(* IEC 61131-3 sources: sis-interlock-demo/src/DUTs/Sis, 21 files *)

(* ---- E_BypassState.dut.st ---- *)
// Назначение: состояние байпаса канала (диаграмма 5.7).
// Автор:      kr0nsch
// Версия:     0.1.0
// Документ:   docs/DESIGN.md, раздел «4.1 Перечисления»
// ВНИМАНИЕ:   код демонстрационный и не предназначен для систем безопасности. Реальная ПАЗ
//             требует определения SIL, сертифицированных аппаратных и программных средств
//             и валидации по ГОСТ Р МЭК 61511.
{attribute 'qualified_only'}
{attribute 'strict'}
TYPE E_BypassState :
(
    Off     := 0,    // байпаса нет
    Active  := 1,    // байпас действует, идёт отсчёт tBypassMax
    Expired := 2,    // срок истёк, запрос ещё держится
    Denied  := 3     // запрос отклонён или байпас снят ключом, запрос ещё держится
) INT;
END_TYPE

(* ---- E_CauseSource.dut.st ---- *)
// Назначение: источник требования причины матрицы: группа голосования или логика приложения
//             (раздел 8.1).
// Автор:      kr0nsch
// Версия:     0.1.0
// Документ:   docs/DESIGN.md, раздел «4.1 Перечисления»
// ВНИМАНИЕ:   код демонстрационный и не предназначен для систем безопасности. Реальная ПАЗ
//             требует определения SIL, сертифицированных аппаратных и программных средств
//             и валидации по ГОСТ Р МЭК 61511.
{attribute 'qualified_only'}
{attribute 'strict'}
TYPE E_CauseSource :
(
    Voting   := 1,   // требование — FB_Voting группы с тем же индексом
    External := 2    // требование — ST_VoteIn.xExtDemand (логика приложения, без голосования)
) INT;
END_TYPE

(* ---- E_ChannelState.dut.st ---- *)
// Назначение: состояние канала группы голосования (таблица 5.1, старшинство: Bypassed, Invalid,
//             Demand, Normal).
// Автор:      kr0nsch
// Версия:     0.1.0
// Документ:   docs/DESIGN.md, раздел «4.1 Перечисления»
// ВНИМАНИЕ:   код демонстрационный и не предназначен для систем безопасности. Реальная ПАЗ
//             требует определения SIL, сертифицированных аппаратных и программных средств
//             и валидации по ГОСТ Р МЭК 61511.
{attribute 'qualified_only'}
{attribute 'strict'}
TYPE E_ChannelState :
(
    NotUsed  := 0,   // канал не входит в схему (номер > N)
    Normal   := 1,   // достоверен, требования нет
    Demand   := 2,   // достоверен, требование срабатывания
    Invalid  := 3,   // недостоверен
    Bypassed := 4    // байпас действует (старше Invalid и Demand)
) INT;
END_TYPE

(* ---- E_DegradePolicy.dut.st ---- *)
// Назначение: политика деградации группы голосования при недостоверных каналах (раздел 5.2).
// Автор:      kr0nsch
// Версия:     0.1.0
// Документ:   docs/DESIGN.md, раздел «4.1 Перечисления»
// ВНИМАНИЕ:   код демонстрационный и не предназначен для систем безопасности. Реальная ПАЗ
//             требует определения SIL, сертифицированных аппаратных и программных средств
//             и валидации по ГОСТ Р МЭК 61511.
{attribute 'qualified_only'}
{attribute 'strict'}
TYPE E_DegradePolicy :
(
    VoteTrip         := 1,   // недостоверный канал голосует «на останов»; 2oo3 → 1oo2 → останов
    DegradeSafe      := 2,   // недостоверный канал исключается, требуется меньше голосов; 2oo3 → 1oo2 → 1oo1
    DegradeAvailable := 3    // недостоверный канал исключается, требуется прежнее число голосов; 2oo3 → 2oo2 → 1oo1
) INT;
END_TYPE

(* ---- E_LimitDir.dut.st ---- *)
// Назначение: направление уставки аналоговой группы голосования (раздел 5.6).
// Автор:      kr0nsch
// Версия:     0.1.0
// Документ:   docs/DESIGN.md, раздел «4.1 Перечисления»
// ВНИМАНИЕ:   код демонстрационный и не предназначен для систем безопасности. Реальная ПАЗ
//             требует определения SIL, сертифицированных аппаратных и программных средств
//             и валидации по ГОСТ Р МЭК 61511.
{attribute 'qualified_only'}
{attribute 'strict'}
TYPE E_LimitDir :
(
    High := 1,       // требование при значении >= уставки
    Low  := 2        // требование при значении <= уставки
) INT;
END_TYPE

(* ---- E_SafeState.dut.st ---- *)
// Назначение: технологический смысл безопасного состояния следствия (для HMI и документов);
//             электрически выход следствия всегда обесточивается (решение D-15).
// Автор:      kr0nsch
// Версия:     0.1.0
// Документ:   docs/DESIGN.md, раздел «4.1 Перечисления»
// ВНИМАНИЕ:   код демонстрационный и не предназначен для систем безопасности. Реальная ПАЗ
//             требует определения SIL, сертифицированных аппаратных и программных средств
//             и валидации по ГОСТ Р МЭК 61511.
{attribute 'qualified_only'}
{attribute 'strict'}
TYPE E_SafeState :
(
    Closed  := 1,    // арматура закрыта
    Open    := 2,    // арматура открыта (сброс давления)
    Stopped := 3,    // механизм остановлен
    Off     := 4,    // потребитель отключён
    Alarm   := 5     // сигнализация включена
) INT;
END_TYPE

(* ---- E_SisEventKind.dut.st ---- *)
// Назначение: коды событий журнала ПАЗ (разделы 4.1, 7.2). В ПЛК нет текстов событий: только
//             коды, индексы и значения (решение D-18).
// Автор:      kr0nsch
// Версия:     0.2.0
// Документ:   docs/DESIGN.md, раздел «4.1 Перечисления»
// ВНИМАНИЕ:   код демонстрационный и не предназначен для систем безопасности. Реальная ПАЗ
//             требует определения SIL, сертифицированных аппаратных и программных средств
//             и валидации по ГОСТ Р МЭК 61511.
{attribute 'qualified_only'}
{attribute 'strict'}
TYPE E_SisEventKind :
(
    None            := 0,    // нет события (пустая запись журнала)
    CauseDemand     := 1,    // требование причины появилось (до задержки)
    CauseClear      := 2,    // требование ушло
    CauseTrip       := 3,    // причина зафиксирована
    FirstOut        := 4,    // первопричина: uiCause = индекс, SIS_FIRST_OUT_START или SIS_FIRST_OUT_CFG
    EffectTrip      := 5,    // следствие обесточено
    EffectRestore   := 6,    // следствие снова под напряжением
    ResetDone       := 7,    // сброс выполнен
    ResetDenied     := 8,    // uiCause — первая мешающая причина или SIS_FIRST_OUT_CFG
    OverrideOn      := 9,    // пусковой обход принят
    OverrideOff     := 10,   // снят командой или ошибкой конфигурации
    OverrideExpired := 11,   // срок обхода истёк или «время назад» (D-19)
    OverrideDenied  := 12,   // запрос обхода отклонён
    BypassOn        := 13,   // байпас канала включён
    BypassOff       := 14,   // снят запросом или ключом разрешения
    BypassExpired   := 15,   // срок байпаса истёк
    BypassDenied    := 16,   // запрос байпаса отклонён
    ChannelInvalid  := 17,   // канал стал недостоверным
    ChannelValid    := 18,   // канал снова достоверен
    DiscrepancyOn   := 19,   // rValue — разброс
    DiscrepancyOff  := 20,   // рассогласование снято
    CfgError        := 21,   // rValue — WORD_TO_REAL(wCfgErr)
    CfgOk           := 22,   // ошибка конфигурации снята
    StartTrip       := 23,   // срабатывание при старте (xStartTripped)
    TimeFault       := 24,   // источник времени пошёл назад: сроки и задержки недостоверны (D-19)
    OverrideCleared := 25    // обход снят автоматически: требования нет непрерывно tOverrideClear (6.4)
) INT;
END_TYPE

(* ---- E_SisInputKind.dut.st ---- *)
// Назначение: вид входов группы голосования: дискретные или аналоговые каналы (раздел 5.6).
// Автор:      kr0nsch
// Версия:     0.1.0
// Документ:   docs/DESIGN.md, раздел «4.1 Перечисления»
// ВНИМАНИЕ:   код демонстрационный и не предназначен для систем безопасности. Реальная ПАЗ
//             требует определения SIL, сертифицированных аппаратных и программных средств
//             и валидации по ГОСТ Р МЭК 61511.
{attribute 'qualified_only'}
{attribute 'strict'}
TYPE E_SisInputKind :
(
    Discrete := 1,   // дискретные каналы axDi / axDiValid
    Analog   := 2    // аналоговые каналы arAi_eu / axAiValid, уставка и гистерезис
) INT;
END_TYPE

(* ---- E_VoteArch.dut.st ---- *)
// Назначение: схема голосования MooN группы каналов (таблица 5.1). ForcedTrip бывает только
//             действующей схемой: голосовать некем или недостоверные каналы уже дают требование.
// Автор:      kr0nsch
// Версия:     0.1.0
// Документ:   docs/DESIGN.md, раздел «4.1 Перечисления»
// ВНИМАНИЕ:   код демонстрационный и не предназначен для систем безопасности. Реальная ПАЗ
//             требует определения SIL, сертифицированных аппаратных и программных средств
//             и валидации по ГОСТ Р МЭК 61511.
{attribute 'qualified_only'}
{attribute 'strict'}
TYPE E_VoteArch :
(
    None       := 0,     // не задана — ошибка конфигурации
    Vote1oo1   := 11,    // один канал
    Vote1oo2   := 12,    // любой из двух
    Vote2oo2   := 22,    // оба из двух
    Vote2oo3   := 23,    // два из трёх
    ForcedTrip := 99     // только действующая схема: голосовать некем или недостоверные каналы уже дают требование
) INT;
END_TYPE

(* ---- ST_CauseCfg.dut.st ---- *)
// Назначение: строка матрицы причин и следствий: включение причины, источник требования,
//             задержка, пусковой обход: срок и подтверждение нормы для автоснятия (раздел 6.4).
// Автор:      kr0nsch
// Версия:     0.2.0
// Документ:   docs/DESIGN.md, раздел «4.2 Структуры»
// ВНИМАНИЕ:   код демонстрационный и не предназначен для систем безопасности. Реальная ПАЗ
//             требует определения SIL, сертифицированных аппаратных и программных средств
//             и валидации по ГОСТ Р МЭК 61511.
{attribute 'qualified_only'}
TYPE ST_CauseCfg :
STRUCT
    xEnable          : BOOL := FALSE;                          // причина используется
    eSource          : E_CauseSource := E_CauseSource.Voting;  // источник требования
    tDelay           : TIME := T#0S;                           // задержка срабатывания, <= SIS_DELAY_MAX
    xOverrideAllowed : BOOL := FALSE;                          // пусковой обход разрешён
    tOverrideMax     : TIME := T#0S;                           // длительность обхода, (0, SIS_OVERRIDE_MAX]
    tOverrideClear   : TIME := T#0S;                           // подтверждение нормы для автоснятия, (0, tOverrideMax)
END_STRUCT
END_TYPE

(* ---- ST_CauseEffectSts.dut.st ---- *)
// Назначение: состояние исполнителя матрицы для HMI, журнала и тестов (раздел 6.3, шаг 8).
// Автор:      kr0nsch
// Версия:     0.2.0
// Документ:   docs/DESIGN.md, раздел «4.2 Структуры»
// ВНИМАНИЕ:   код демонстрационный и не предназначен для систем безопасности. Реальная ПАЗ
//             требует определения SIL, сертифицированных аппаратных и программных средств
//             и валидации по ГОСТ Р МЭК 61511.
{attribute 'qualified_only'}
TYPE ST_CauseEffectSts :
STRUCT
    uiFirstOut       : UINT;        // SIS_FIRST_OUT_NONE, 1..N, SIS_FIRST_OUT_START или SIS_FIRST_OUT_CFG
    ltFirstOut       : LTIME;       // момент фиксации первопричины (I_TimeSource); LTIME#0S — нет
    wFirstOutMask    : WORD;        // все причины, зафиксированные в вызове первопричины
    wCausePresent    : WORD;        // требование есть сейчас (до задержки), причина включена
    wCauseActive     : WORD;        // требование после задержки (без учёта обхода)
    wCauseLatched    : WORD;        // причина зафиксирована, до сброса
    wOverridden      : WORD;        // пусковой обход действует
    wEffectTripped   : WORD;        // следствие сработало (выход обесточен), j <= uiEffectCount
    xTripped         : BOOL;        // хотя бы одно следствие сработало
    xResetPermitted  : BOOL;        // сброс сейчас разрешён
    uiResetBlocker   : UINT;        // 0 — нет; первая мешающая причина; SIS_FIRST_OUT_CFG — ошибка конфигурации
    xCfgError        : BOOL;        // ошибка конфигурации матрицы
    wCfgErr          : WORD;        // биты CEM_CFG_*
    udiTripCount     : UDINT;       // фиксаций первопричины с запуска
    atOverrideRemain : ARRAY[1..GVL_Const.SIS_CAUSES_MAX] OF TIME;   // остаток обхода; T#0S — обхода нет
    atDelayRemain    : ARRAY[1..GVL_Const.SIS_CAUSES_MAX] OF TIME;   // остаток задержки; T#0S — отсчёта нет
    // остаток подтверждения нормы до автоснятия обхода (6.4, п. 5); T#0S — обхода нет или требование есть
    atOverrideClearRemain : ARRAY[1..GVL_Const.SIS_CAUSES_MAX] OF TIME;
END_STRUCT
END_TYPE

(* ---- ST_CemCfg.dut.st ---- *)
// Назначение: конфигурация матрицы причин и следствий с CRC. Значения по умолчанию дают ошибку
//             конфигурации (uiCauseCount = 0) — срабатывание всех следствий (раздел 6.8).
// Автор:      kr0nsch
// Версия:     0.1.0
// Документ:   docs/DESIGN.md, раздел «4.2 Структуры»
// ВНИМАНИЕ:   код демонстрационный и не предназначен для систем безопасности. Реальная ПАЗ
//             требует определения SIL, сертифицированных аппаратных и программных средств
//             и валидации по ГОСТ Р МЭК 61511.
{attribute 'qualified_only'}
TYPE ST_CemCfg :
STRUCT
    uiCauseCount  : UINT := 0;      // используемых причин, 1..SIS_CAUSES_MAX; 0 — ошибка (fail-safe)
    uiEffectCount : UINT := 0;      // используемых следствий, 1..SIS_EFFECTS_MAX
    xStartTripped : BOOL := TRUE;   // после старта ПЛК все следствия сработали до первого сброса
    astCause      : ARRAY[1..GVL_Const.SIS_CAUSES_MAX] OF ST_CauseCfg;     // строки матрицы
    astEffect     : ARRAY[1..GVL_Const.SIS_EFFECTS_MAX] OF ST_EffectCfg;   // столбцы матрицы
    wMatrixCrc    : WORD := 0;      // CRC-16/CCITT-FALSE матрицы (раздел 6.8), считает генератор
END_STRUCT
END_TYPE

(* ---- ST_CemCmd.dut.st ---- *)
// Назначение: импульсные команды HMI исполнителю матрицы; FB_CauseEffect сбрасывает их в том же
//             вызове (разделы 6.4, 6.5).
// Автор:      kr0nsch
// Версия:     0.1.0
// Документ:   docs/DESIGN.md, раздел «4.2 Структуры»
// ВНИМАНИЕ:   код демонстрационный и не предназначен для систем безопасности. Реальная ПАЗ
//             требует определения SIL, сертифицированных аппаратных и программных средств
//             и валидации по ГОСТ Р МЭК 61511.
{attribute 'qualified_only'}
TYPE ST_CemCmd :
STRUCT
    xReset           : BOOL;        // сброс ПАЗ
    xStartupOverride : BOOL;        // пусковой обход всех причин с xOverrideAllowed
    wOverrideReq     : WORD;        // обход причин по маске
    wOverrideCancel  : WORD;        // снять обход по маске
END_STRUCT
END_TYPE

(* ---- ST_EffectCfg.dut.st ---- *)
// Назначение: столбец матрицы причин и следствий: смысл безопасного состояния и маска причин,
//             которые отключают следствие (раздел 6.7).
// Автор:      kr0nsch
// Версия:     0.1.0
// Документ:   docs/DESIGN.md, раздел «4.2 Структуры»
// ВНИМАНИЕ:   код демонстрационный и не предназначен для систем безопасности. Реальная ПАЗ
//             требует определения SIL, сертифицированных аппаратных и программных средств
//             и валидации по ГОСТ Р МЭК 61511.
{attribute 'qualified_only'}
TYPE ST_EffectCfg :
STRUCT
    eSafeState : E_SafeState := E_SafeState.Off;   // смысл для HMI и документов; выход всегда обесточивается
    wCauseMask : WORD := 0;                        // бит i-1 — причина i отключает это следствие («X» в столбце)
END_STRUCT
END_TYPE

(* ---- ST_SisCmd.dut.st ---- *)
// Назначение: команды HMI узлу ПАЗ: матрица и байпасы каналов по причинам (раздел 8.1).
// Автор:      kr0nsch
// Версия:     0.1.0
// Документ:   docs/DESIGN.md, раздел «4.2 Структуры»
// ВНИМАНИЕ:   код демонстрационный и не предназначен для систем безопасности. Реальная ПАЗ
//             требует определения SIL, сертифицированных аппаратных и программных средств
//             и валидации по ГОСТ Р МЭК 61511.
{attribute 'qualified_only'}
TYPE ST_SisCmd :
STRUCT
    stCem   : ST_CemCmd;                                          // сброс и пусковые обходы
    astVote : ARRAY[1..GVL_Const.SIS_CAUSES_MAX] OF ST_VoteCmd;   // байпасы каналов по причинам
END_STRUCT
END_TYPE

(* ---- ST_SisEvent.dut.st ---- *)
// Назначение: запись журнала событий ПАЗ. Порядок полей — без выравнивающих пропусков:
//             SIZEOF = 24 байта (раздел 4.2, тест Log_SizeOfEvent_Is24).
// Автор:      kr0nsch
// Версия:     0.1.0
// Документ:   docs/DESIGN.md, раздел «4.2 Структуры»
// ВНИМАНИЕ:   код демонстрационный и не предназначен для систем безопасности. Реальная ПАЗ
//             требует определения SIL, сертифицированных аппаратных и программных средств
//             и валидации по ГОСТ Р МЭК 61511.
{attribute 'qualified_only'}
TYPE ST_SisEvent :
STRUCT
    ltTime    : LTIME;              // монотонная отметка источника времени
    udiSeq    : UDINT;              // номер события; присваивает журнал (1, 2, ...; после 16#FFFFFFFF — 1)
    rValue    : REAL;               // значение канала, разброс, код ошибки; иначе 0.0
    eKind     : E_SisEventKind;     // вид события
    uiCause   : UINT;               // 0 — нет; 1..N; SIS_FIRST_OUT_START / SIS_FIRST_OUT_CFG
    uiEffect  : UINT;               // 0 — нет; 1..M
    uiChannel : UINT;               // 0 — нет; 1..3
END_STRUCT
END_TYPE

(* ---- ST_VoteCmd.dut.st ---- *)
// Назначение: команды группы голосования от HMI — уровни: запрос байпаса держится, пока нужен;
//             FB_Voting их не сбрасывает (раздел 5.7).
// Автор:      kr0nsch
// Версия:     0.1.0
// Документ:   docs/DESIGN.md, раздел «4.2 Структуры»
// ВНИМАНИЕ:   код демонстрационный и не предназначен для систем безопасности. Реальная ПАЗ
//             требует определения SIL, сертифицированных аппаратных и программных средств
//             и валидации по ГОСТ Р МЭК 61511.
{attribute 'qualified_only'}
TYPE ST_VoteCmd :
STRUCT
    axBypassReq : ARRAY[1..GVL_Const.SIS_VOTE_CH_MAX] OF BOOL;  // запрос байпаса канала (держится, пока нужен)
END_STRUCT
END_TYPE

(* ---- ST_VoteIn.dut.st ---- *)
// Назначение: сигналы каналов одной группы голосования: дискретные значения с контролем линии,
//             аналоговые значения в инж. ед. с достоверностью, внешнее требование (раздел 5.6).
// Автор:      kr0nsch
// Версия:     0.1.0
// Документ:   docs/DESIGN.md, раздел «4.2 Структуры»
// ВНИМАНИЕ:   код демонстрационный и не предназначен для систем безопасности. Реальная ПАЗ
//             требует определения SIL, сертифицированных аппаратных и программных средств
//             и валидации по ГОСТ Р МЭК 61511.
{attribute 'qualified_only'}
TYPE ST_VoteIn :
STRUCT
    axDi       : ARRAY[1..GVL_Const.SIS_VOTE_CH_MAX] OF BOOL;   // дискретные каналы (значение с поля)
    axDiValid  : ARRAY[1..GVL_Const.SIS_VOTE_CH_MAX] OF BOOL;   // контроль линии / диагностика: TRUE — исправен
    arAi_eu    : ARRAY[1..GVL_Const.SIS_VOTE_CH_MAX] OF REAL;   // аналоговые каналы, инж. ед.
    axAiValid  : ARRAY[1..GVL_Const.SIS_VOTE_CH_MAX] OF BOOL;   // достоверность (NE 43 и т. п.): TRUE — достоверен
    xExtDemand : BOOL;                                          // для eSource = External: TRUE — требование
END_STRUCT
END_TYPE

(* ---- ST_VoteResult.dut.st ---- *)
// Назначение: результат F_VoteEval: требование, деградация, действующая схема и счётчики
//             состояний каналов (раздел 5.2).
// Автор:      kr0nsch
// Версия:     0.1.0
// Документ:   docs/DESIGN.md, раздел «4.2 Структуры»
// ВНИМАНИЕ:   код демонстрационный и не предназначен для систем безопасности. Реальная ПАЗ
//             требует определения SIL, сертифицированных аппаратных и программных средств
//             и валидации по ГОСТ Р МЭК 61511.
{attribute 'qualified_only'}
TYPE ST_VoteResult :
STRUCT
    xTrip      : BOOL := TRUE;                      // TRUE — требование срабатывания
    xDegraded  : BOOL;                              // есть байпасированные или недостоверные каналы
    eArchEff   : E_VoteArch := E_VoteArch.None;     // действующая схема
    uiDemand   : UINT;                              // каналов Demand
    uiInvalid  : UINT;                              // каналов Invalid
    uiBypassed : UINT;                              // каналов Bypassed
    uiNormal   : UINT;                              // каналов Normal
END_STRUCT
END_TYPE

(* ---- ST_VotingCfg.dut.st ---- *)
// Назначение: конфигурация группы голосования. Значения по умолчанию дают ошибку конфигурации
//             (eArch = None) — срабатывание группы (fail-safe, раздел 3.4).
// Автор:      kr0nsch
// Версия:     0.1.0
// Документ:   docs/DESIGN.md, раздел «4.2 Структуры»
// ВНИМАНИЕ:   код демонстрационный и не предназначен для систем безопасности. Реальная ПАЗ
//             требует определения SIL, сертифицированных аппаратных и программных средств
//             и валидации по ГОСТ Р МЭК 61511.
{attribute 'qualified_only'}
TYPE ST_VotingCfg :
STRUCT
    eArch              : E_VoteArch := E_VoteArch.None;                  // None — ошибка (fail-safe)
    ePolicy            : E_DegradePolicy := E_DegradePolicy.VoteTrip;    // политика деградации
    eInput             : E_SisInputKind := E_SisInputKind.Discrete;      // вид входов
    xDiHealthy         : BOOL := TRUE;     // значение дискретного канала в норме; другое — требование
    eLimitDir          : E_LimitDir := E_LimitDir.High;                  // направление уставки (Analog)
    rTripLimit_eu      : REAL := 0.0;      // уставка срабатывания, инж. ед. (включительно)
    rHyst_eu           : REAL := 0.0;      // гистерезис снятия требования, >= 0
    rDiscrepancyMax_eu : REAL := 0.0;      // допустимый разброс каналов; 0.0 — контроль выключен
    tDiscrepancyDelay  : TIME := T#0S;     // задержка тревоги рассогласования
    tBypassMax         : TIME := T#0S;     // максимальная длительность байпаса; T#0S — байпас запрещён
    uiMaxBypass        : UINT := 0;        // одновременных байпасов в группе, 0..N-1
END_STRUCT
END_TYPE

(* ---- ST_VotingSts.dut.st ---- *)
// Назначение: состояние группы голосования для HMI, журнала и тестов (раздел 5.5, шаг 9).
// Автор:      kr0nsch
// Версия:     0.1.0
// Документ:   docs/DESIGN.md, раздел «4.2 Структуры»
// ВНИМАНИЕ:   код демонстрационный и не предназначен для систем безопасности. Реальная ПАЗ
//             требует определения SIL, сертифицированных аппаратных и программных средств
//             и валидации по ГОСТ Р МЭК 61511.
{attribute 'qualified_only'}
TYPE ST_VotingSts :
STRUCT
    xTrip          : BOOL := TRUE;                  // TRUE — требование срабатывания (= FB_Voting.xTrip)
    eArchEff       : E_VoteArch := E_VoteArch.None; // действующая схема
    xDegraded      : BOOL;            // есть байпасированные или недостоверные каналы
    xCfgError      : BOOL;            // ошибка конфигурации группы
    wCfgErr        : WORD;            // биты VOTE_CFG_*
    xDiscrepancy   : BOOL;            // тревога рассогласования (после задержки)
    rSpread_eu     : REAL;            // max − min участвующих аналоговых каналов; 0.0, если их меньше двух
    uiDemand       : UINT;            // каналов Demand
    uiInvalid      : UINT;            // каналов Invalid
    uiBypassed     : UINT;            // каналов Bypassed
    uiNormal       : UINT;            // каналов Normal
    aeChState      : ARRAY[1..GVL_Const.SIS_VOTE_CH_MAX] OF E_ChannelState;   // состояния каналов
    aeBypass       : ARRAY[1..GVL_Const.SIS_VOTE_CH_MAX] OF E_BypassState;    // состояния байпасов
    atBypassRemain : ARRAY[1..GVL_Const.SIS_VOTE_CH_MAX] OF TIME;   // остаток байпаса; T#0S, если не Active
END_STRUCT
END_TYPE
